// TIA Portal V17 export
// export: Created 2026-11-17T10:42:13.4013486Z, ExportSetting WithDefaults, DisplayName Totally Integrated Automation Portal, DisplayVersion V17, DisplayName TIA Portal Openness, DisplayVersion V17, DisplayName TIA Portal Version Control Interface, DisplayVersion V17, DisplayName STEP 7 Professional, DisplayVersion V17, DisplayName STEP 7 Safety, DisplayVersion V17, DisplayName WinCC Advanced, DisplayVersion V17
TagTable "红绿灯HMI变量"
  StartPB : Bool  (PLC tag StartPB, HMI_连接_1, 100 ms)
  StopPB : Bool  (PLC tag StopPB, HMI_连接_1, 100 ms)
  Run : Bool  (PLC tag Run, HMI_连接_1, 100 ms)
  NS_Red : Bool  (PLC tag NS_Red, HMI_连接_1, 100 ms)
  NS_Yellow : Bool  (PLC tag NS_Yellow, HMI_连接_1, 100 ms)
  NS_Green : Bool  (PLC tag NS_Green, HMI_连接_1, 100 ms)
  EW_Red : Bool  (PLC tag EW_Red, HMI_连接_1, 100 ms)
  EW_Yellow : Bool  (PLC tag EW_Yellow, HMI_连接_1, 100 ms)
  EW_Green : Bool  (PLC tag EW_Green, HMI_连接_1, 100 ms)
